// TIA Portal V19 export
// export: Created 2026-10-15T09:44:24.9257696Z, ExportSetting WithDefaults, DisplayName Totally Integrated Automation Portal, DisplayVersion V19, DisplayName TIA Portal Openness, DisplayVersion V19, DisplayName TIA Portal Version Control Interface, DisplayVersion V19, DisplayName STEP 7 Professional, DisplayVersion V19, DisplayName STEP 7 Safety, DisplayVersion V19, DisplayName WinCC Basic/Comfort/Advanced, DisplayVersion V19, DisplayName WinCC Unified, DisplayVersion V19
FUNCTION "ROLL_PB25" : Void   // FC32, SCL
{ S7_Optimized_Access := 'TRUE' }
VERSION : 0.1
// stored: AutoNumber true, IsIECCheckEnabled false, SetENOAutomatically false, UDAEnableTagReadback false
   VAR_TEMP
      r : Bool;
      a1 : Word;
      a2 : Word;
      activeDataBlock : Int;
      comparisonResults : Array[0..14] of Bool;
   END_VAR
BEGIN

   #r := FALSE;
   #a1 := W#16#0000;
   #a2 := W#16#0000;
   #activeDataBlock := 0;
   // PB25, STEP 5 network 1
   #activeDataBlock := 15;
   // PB25, STEP 5 network 2
   #a2 := #a1;
   #a1 := "ROLL_GetM"(FirstByte := 5, Width := 8);
   #a2 := #a1;
   #a1 := W#16#0000;
   #comparisonResults[0] := (WORD_TO_INT(#a2) <> WORD_TO_INT(#a1));
   #r := #comparisonResults[0];
   "ROLL_State".M[87, 0] := #r;
   // PB25, STEP 5 network 3
   #a2 := #a1;
   #a1 := "ROLL_GetM"(FirstByte := 6, Width := 8);
   #a2 := #a1;
   #a1 := W#16#0000;
   #comparisonResults[1] := (WORD_TO_INT(#a2) <> WORD_TO_INT(#a1));
   #r := #comparisonResults[1];
   "ROLL_State".M[87, 1] := #r;
   // PB25, STEP 5 network 4
   #a2 := #a1;
   #a1 := "ROLL_GetM"(FirstByte := 7, Width := 8);
   #a2 := #a1;
   #a1 := W#16#0000;
   #comparisonResults[2] := (WORD_TO_INT(#a2) <> WORD_TO_INT(#a1));
   #r := #comparisonResults[2];
   "ROLL_State".M[87, 2] := #r;
   // PB25, STEP 5 network 5
   #a2 := #a1;
   #a1 := "ROLL_GetM"(FirstByte := 8, Width := 8);
   #a2 := #a1;
   #a1 := W#16#0000;
   #comparisonResults[3] := (WORD_TO_INT(#a2) <> WORD_TO_INT(#a1));
   #r := #comparisonResults[3];
   "ROLL_State".M[87, 3] := #r;
   // PB25, STEP 5 network 6
   #a2 := #a1;
   #a1 := "ROLL_GetM"(FirstByte := 9, Width := 8);
   #a2 := #a1;
   #a1 := W#16#0000;
   #comparisonResults[4] := (WORD_TO_INT(#a2) <> WORD_TO_INT(#a1));
   #r := #comparisonResults[4];
   "ROLL_State".M[87, 4] := #r;
   // PB25, STEP 5 network 7
   #a2 := #a1;
   #a1 := "ROLL_GetM"(FirstByte := 10, Width := 8);
   #a2 := #a1;
   #a1 := W#16#0000;
   #comparisonResults[5] := (WORD_TO_INT(#a2) <> WORD_TO_INT(#a1));
   #r := #comparisonResults[5];
   "ROLL_State".M[87, 5] := #r;
   // PB25, STEP 5 network 8
   #a2 := #a1;
   #a1 := "ROLL_GetM"(FirstByte := 11, Width := 8);
   #a2 := #a1;
   #a1 := W#16#0000;
   #comparisonResults[6] := (WORD_TO_INT(#a2) <> WORD_TO_INT(#a1));
   #r := #comparisonResults[6];
   "ROLL_State".M[87, 6] := #r;
   // PB25, STEP 5 network 9
   #a2 := #a1;
   #a1 := "ROLL_GetM"(FirstByte := 12, Width := 8);
   #a2 := #a1;
   #a1 := W#16#0000;
   #comparisonResults[7] := (WORD_TO_INT(#a2) <> WORD_TO_INT(#a1));
   #r := #comparisonResults[7];
   "ROLL_State".M[87, 7] := #r;
   // PB25, STEP 5 network 10
   #a2 := #a1;
   #a1 := "ROLL_GetM"(FirstByte := 13, Width := 8);
   #a2 := #a1;
   #a1 := W#16#0000;
   #comparisonResults[8] := (WORD_TO_INT(#a2) <> WORD_TO_INT(#a1));
   #r := #comparisonResults[8];
   "ROLL_State".M[88, 0] := #r;
   // PB25, STEP 5 network 11
   #a2 := #a1;
   #a1 := "ROLL_GetM"(FirstByte := 14, Width := 8);
   #a2 := #a1;
   #a1 := W#16#0000;
   #comparisonResults[9] := (WORD_TO_INT(#a2) <> WORD_TO_INT(#a1));
   #r := #comparisonResults[9];
   "ROLL_State".M[88, 1] := #r;
   // PB25, STEP 5 network 12
   #a2 := #a1;
   #a1 := "ROLL_GetM"(FirstByte := 15, Width := 8);
   #a2 := #a1;
   #a1 := W#16#0000;
   #comparisonResults[10] := (WORD_TO_INT(#a2) <> WORD_TO_INT(#a1));
   #r := #comparisonResults[10];
   "ROLL_State".M[88, 2] := #r;
   // PB25, STEP 5 network 13
   #a2 := #a1;
   #a1 := "ROLL_GetM"(FirstByte := 16, Width := 8);
   #a2 := #a1;
   #a1 := W#16#0000;
   #comparisonResults[11] := (WORD_TO_INT(#a2) <> WORD_TO_INT(#a1));
   #r := #comparisonResults[11];
   "ROLL_State".M[88, 3] := #r;
   // PB25, STEP 5 network 14
   #a2 := #a1;
   #a1 := "ROLL_GetM"(FirstByte := 17, Width := 8);
   #a2 := #a1;
   #a1 := W#16#0000;
   #comparisonResults[12] := (WORD_TO_INT(#a2) <> WORD_TO_INT(#a1));
   #r := #comparisonResults[12];
   "ROLL_State".M[88, 4] := #r;
   // PB25, STEP 5 network 15
   #a2 := #a1;
   #a1 := "ROLL_GetM"(FirstByte := 18, Width := 8);
   #a2 := #a1;
   #a1 := W#16#0000;
   #comparisonResults[13] := (WORD_TO_INT(#a2) <> WORD_TO_INT(#a1));
   #r := #comparisonResults[13];
   "ROLL_State".M[88, 5] := #r;
   // PB25, STEP 5 network 16
   #a2 := #a1;
   #a1 := "ROLL_GetM"(FirstByte := 19, Width := 8);
   #a2 := #a1;
   #a1 := W#16#0000;
   #comparisonResults[14] := (WORD_TO_INT(#a2) <> WORD_TO_INT(#a1));
   #r := #comparisonResults[14];
   "ROLL_State".M[88, 6] := #r;
   // PB25, STEP 5 network 17
   #r := ("ROLL_State".M[87, 0] OR "ROLL_State".M[87, 1] OR "ROLL_State".M[87, 2] OR "ROLL_State".M[87, 3] OR "ROLL_State".M[87, 4] OR "ROLL_State".M[87, 5] OR "ROLL_State".M[87, 6] OR "ROLL_State".M[87, 7] OR "ROLL_State".M[88, 0] OR "ROLL_State".M[88, 1] OR "ROLL_State".M[88, 2] OR "ROLL_State".M[88, 3] OR "ROLL_State".M[88, 4] OR "ROLL_State".M[88, 5] OR "ROLL_State".M[88, 6]);
   "ROLL_State".M[88, 7] := #r;
   // PB25, STEP 5 network 18
   #r := ("ROLL_IO".Input[1, 2] OR "ROLL_State".M[88, 7]);
   "ROLL_IO".Output[16, 4] := #r;
   // PB25, STEP 5 network 19
   #r := (("ROLL_State".M[3, 6] AND "ROLL_State".M[31, 6]) OR "ROLL_IO".Input[1, 2]);
   "ROLL_IO".Output[16, 5] := #r;
   // PB25, STEP 5 network 20
   #r := ("ROLL_IO".Input[1, 2] OR "ROLL_IO".Input[3, 4]);
   "ROLL_IO".Output[16, 0] := #r;
   // PB25, STEP 5 network 21
   #r := (((NOT "ROLL_State".M[31, 5]) AND "ROLL_State".M[28, 4]) OR ("ROLL_State".M[3, 6] AND "ROLL_State".M[74, 0]) OR "ROLL_IO".Input[1, 2]);
   "ROLL_IO".Output[16, 2] := #r;
   // PB25, STEP 5 network 22
   #r := (("ROLL_State".M[3, 6] AND "ROLL_State".M[31, 5]) OR "ROLL_IO".Input[1, 2] OR "ROLL_State".M[31, 4]);
   "ROLL_IO".Output[16, 3] := #r;
   // PB25, STEP 5 network 23
   #r := "ROLL_IO".Input[2, 0];
   "ROLL_IO".Output[19, 3] := #r;
   // PB25, STEP 5 network 24
   #r := (((("ROLL_IO".Input[14, 0] AND "ROLL_State".M[37, 1]) OR "ROLL_State".M[53, 6]) AND "ROLL_IO".Input[0, 2]) OR ("ROLL_IO".Input[0, 1] AND "ROLL_State".M[190, 6] AND "ROLL_State".M[20, 7]));
   IF #r THEN
       "ROLL_State".M[71, 5] := TRUE;
   END_IF;
   #r := (("ROLL_IO".Input[0, 1] AND "ROLL_State".M[190, 5] AND "ROLL_State".M[20, 7]) OR ("ROLL_IO".Input[0, 2] AND "ROLL_State".M[37, 2]));
   IF #r THEN
       "ROLL_State".M[71, 5] := FALSE;
   END_IF;
   #r := "ROLL_State".M[71, 5];
   "ROLL_IO".Output[17, 7] := #r;
   // PB25, STEP 5 network 25
   RETURN;
END_FUNCTION
